(* IEC 61131-3 sources: PLC-Static-Analysis/modules/plc-rules/src/test/resources/PLCA-P004/notasks, 1 file *)

(* ---- two.st ---- *)
VAR_GLOBAL
    gnParts : INT;
END_VAR

PROGRAM P_A
gnParts := 1;
END_PROGRAM

PROGRAM P_B
gnParts := 2;
END_PROGRAM
